// TIA Portal V19 export
TYPE "AnaMon.Permission"
   STRUCT
      MsgSupEn : Bool;
      HiAlmSupEn : Bool;
      HiWrnSupEn : Bool;
      LoWrnSupEn : Bool;
      LoAlmSupEn : Bool;
   END_STRUCT;
END_TYPE
